Fanuc KAREL source: kt00908.KL

-- PROVISIONAL review KL for V770-1; original PC SHA256 411b5863faf1b006ef806257a9ae76e56cd8974e0067a145549089de90dfe52c
-- Incomplete behavior may be omitted. Consult companion uncertainty JSON. Do not deploy.
PROGRAM KT00908
%NOLOCKGROUP
BEGIN
  -- UNRESOLVED_PC offsets 5-28; opcodes 27,22,1C,31,4A
  -- UNRESOLVED_PC offsets 33-37; opcodes 7F
END KT00908
